Fanuc KAREL source: KD00069.KL

PROGRAM KD00069
%NOLOCKGROUP
VAR
  I: INTEGER
  J: INTEGER
  B: BOOLEAN
  R: REAL
  S: STRING[80]
BEGIN
  CONDITION[1]:
  WHEN DIN[1] = ON DO
    RESUME
  ENDCONDITION
END KD00069
